(* IEC 61131-3 sources: PLC_Gen_Frame/Agents4PLC_release/results/task_1e189b8d, 1 file *)

(* ---- output.ST ---- *)
FUNCTION_BLOCK CottonCandyMachine
VAR_INPUT
    SugarLevel : REAL; (* Input for sugar level *)
    SpinningSpeed : INT; (* Input for spinning speed *)
END_VAR
VAR_OUTPUT
    SugarFeeder : BOOL; (* Output to control sugar feeding *)
    MotorSpeed : INT; (* Output to control spinning motor speed *)
END_VAR

// Control sugar feeder activation based on sugar level threshold
SugarFeeder := SugarLevel < 10.0;

// Set motor speed to input value if positive, otherwise set to 0
IF SpinningSpeed > 0 THEN
    MotorSpeed := SpinningSpeed;
ELSE
    MotorSpeed := 0;
END_IF;

END_FUNCTION_BLOCK
